FUNCTION_BLOCK PARTS_COUNTER (* Migrated from IEC 61131-3 ST *)
  (* Standard: 61499-2 *)
  (* Version 1.0, 2026-11-06, st2fb *)
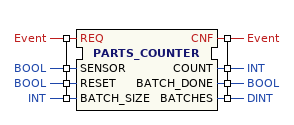
  EVENT_INPUT
    REQ WITH SENSOR, RESET, BATCH_SIZE;
  END_EVENT
  EVENT_OUTPUT
    CNF WITH COUNT, BATCH_DONE, BATCHES;
  END_EVENT
  VAR_INPUT
    SENSOR : BOOL;
    RESET : BOOL;
    BATCH_SIZE : INT;
  END_VAR
  VAR_OUTPUT
    COUNT : INT;
    BATCH_DONE : BOOL;
    BATCHES : DINT;
  END_VAR
  VAR
    COUNTER_CU : BOOL := FALSE;
    COUNTER_R : BOOL := FALSE;
    COUNTER_PV : INT := 0;
    COUNTER_Q : BOOL := FALSE;
    COUNTER_CV : INT := 0;
    COUNTER_CU_T_Q : BOOL := FALSE;
    COUNTER_CU_T_M : BOOL := FALSE;
    DONE_EDGE_CLK : BOOL := FALSE;
    DONE_EDGE_Q : BOOL := FALSE;
    DONE_EDGE_M : BOOL := FALSE;
  END_VAR
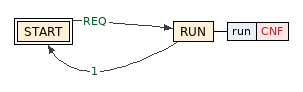
  EC_STATES
    START;
    RUN : run -> CNF;
  END_STATES
  EC_TRANSITIONS
    START TO RUN := REQ;
    RUN TO START := 1;
  END_TRANSITIONS
  ALGORITHM run IN ST:
COUNTER_CU := SENSOR;
COUNTER_R := RESET OR DONE_EDGE_Q;
COUNTER_PV := BATCH_SIZE;
COUNTER_CU_T_Q := COUNTER_CU AND NOT COUNTER_CU_T_M;
COUNTER_CU_T_M := COUNTER_CU;
IF COUNTER_R THEN
  COUNTER_CV := 0;
ELSIF COUNTER_CU_T_Q AND (COUNTER_CV < COUNTER_PV) THEN
  COUNTER_CV := COUNTER_CV + 1;
END_IF;
COUNTER_Q := COUNTER_CV >= COUNTER_PV;
COUNT := COUNTER_CV;
BATCH_DONE := COUNTER_Q;
DONE_EDGE_CLK := COUNTER_Q;
DONE_EDGE_Q := DONE_EDGE_CLK AND NOT DONE_EDGE_M;
DONE_EDGE_M := DONE_EDGE_CLK;
IF DONE_EDGE_Q THEN
  BATCHES := BATCHES + 1;
END_IF;
IF RESET THEN
  BATCHES := 0;
END_IF;
  END_ALGORITHM
END_FUNCTION_BLOCK
